// TIA Portal V20 export
// export: Created 2026-10-20T12:45:28.6356782Z, ExportSetting WithDefaults, DisplayName Totally Integrated Automation Portal, DisplayVersion V20 Update 6, DisplayName TIA Portal Openness, DisplayVersion V20 Update 6, DisplayName TIA Portal Version Control Interface, DisplayVersion V20 Update 6, DisplayName SINAMICS Startdrive Advanced, DisplayVersion V20 SP1, DisplayName SINAMICS Startdrive G130, G150, S120, S150, SINAMICS MV, G220, S200, S210, DisplayVersion V20 SP1, DisplayName SINAMICS Startdrive G110M, G120, G120C, G120D, G120P, G115D, DisplayVersion V20 SP1, DisplayName STEP 7 Professional, DisplayVersion V20 Update 6, DisplayName STEP 7 Safety, DisplayVersion V20 Update 2, DisplayName WinCC Basic/Comfort/Advanced, DisplayVersion V20 Update 6, DisplayName WinCC Unified, DisplayVersion V20 Update 6
DATA_BLOCK "VTD_HMI_FB_2_DB"   // DB60
VERSION : 0.1
// stored: AutoNumber true, DBAccessibleFromOPCUA true, InstanceOfName VTD_HMI_FB_1, InstanceOfType FB
"VTD_HMI_FB_1"
   // VAR_INPUT
   //    HMI_No : UInt;
   //    HMI_Box { ExternalAccessible := 'False'; ExternalVisible := 'False'; ExternalWritable := 'False'} : UInt;
   //    Sys_No : UInt;
   // END_VAR
   // VAR
   //    T_Charge { S7_SetPoint := 'True'} : TON_TIME;
   //    T_Charge_IN : Bool;
   //    Charged : Bool;
   // END_VAR
BEGIN
END_DATA_BLOCK
